Staubli VAL3: click_logExport.pgx

program click_logExport()
  local num l_nResult
  local string l_sDate
begin
  l_sDate=getDate("%m_%d %H_%M_%S")
  call rs:saveLog("USB0://LOG_"+l_sDate+"/log",l_nResult)
  if l_nResult!=0
    call rs:saveLog("SP2_USB0://LOG_"+l_sDate+"/log",l_nResult)
    if l_nResult!=0
      popUpMsg("未识别U盘,导出失败:"+toString("",l_nResult))
      return
    endIf
  endIf
  popUpMsg("导出到U盘成功,文件名:LOG_"+l_sDate)
end
